Yaskawa INFORM job: LONGPRO3.JBI

/JOB
//NAME LONGPRO3
//POS
///NPOS 4,0,4,0,0,0
///TOOL 9
///POSTYPE PULSE
///PULSE
C00000=0,0,0
C00001=0,0,0
C00002=0,0,0
C00003=0,0,0
EC00000=0
EC00001=0
EC00002=0
EC00003=0
//INST
<volatile>
///COMM Generated using RoboDK
///ATTR SC,RW
///GROUP1 RB1
NOP
'10.0,20.0,150.0,0.0,0.0,0.0
MOVJ C00000 VJ=50.00  +MOVJ EC00000 VJ=100.00
MOVJ C00001 VJ=50.00  +MOVJ EC00001 VJ=100.00
MOVJ C00002 VJ=50.00  +MOVJ EC00002 VJ=100.00
MOVJ C00003 VJ=50.00  +MOVJ EC00003 VJ=100.00
END
